(* IEC 61131-3 sources: daoli-st-library/_quarantine/R80, 3 files *)

(* ---- FC_DL_HydroPipePressDrop.st ---- *)
(*
  ============================================================
  组件名 : FC_DL_HydroPipePressDrop
  分类   : DL_Device
  功能   : 液压管路压降计算，由流量管径长度求流速、雷诺数、摩阻系数与压降
  开源溯源 : internal-design（本轮无外部代码逐行引用）
             参考语义 : 无外部参考
  复杂度 : C2
  版本   : 1.0.0
  ============================================================
  口径说明 : 工作介质取液压油，密度按 850 kg/m3 常量代入；黏度由 cSt 折算为 m2/s；
             层流区用 64/Re，湍流区用 Blasius 式 0.3164/Re^0.25；粗糙度引脚仅登记
             供上层记录，本件不进入摩阻判据（Colebrook 迭代属另一件边界）。
*)

FUNCTION FC_DL_HydroPipePressDrop : REAL
VAR_INPUT
    rFlow_lpm  : REAL; // 体积流量 [l/min] volume flow [l per minute]
    rDia_mm    : REAL; // 管内径 [mm] pipe inner diameter [mm]
    rLength_m  : REAL; // 管长 [m] pipe length [m]
    rVisc_cSt  : REAL; // 运动黏度 [cSt] kinematic viscosity [centistoke]
    rRough_mm  : REAL; // 管内壁粗糙度 [mm] inner wall roughness [mm]
END_VAR
VAR_OUTPUT
    rVel_m_s : REAL; // 管内流速 [m/s] pipe velocity [m per second]
    rRe      : REAL; // 雷诺数 [无量纲] Reynolds number [dimensionless]
    rDrop_bar: REAL; // 沿程压降 [bar] friction pressure drop [bar]
    bValid   : BOOL; // 结果有效标志 result validity flag
END_VAR
VAR CONSTANT
    DL_PI_4     : REAL := 0.7853982; // 四分之圆周率 pi divided by four
    DL_MM_TO_M  : REAL := 1000.0; // 每米毫米数 millimetres per metre
    DL_LPM_TO_M3S : REAL := 60000.0; // 升每分到立方米每秒的除数 divisor from litre per minute to cubic metre per second
    DL_CST_TO_M2S : REAL := 1.0E-6; // 厘斯到平方米每秒的乘子 multiplier from centistoke to square metre per second
    DL_DENSITY  : REAL := 850.0; // 液压油密度 [kg/m3] hydraulic oil density [kg per cubic metre]
    DL_RE_LAM   : REAL := 2300.0; // 层流上限雷诺数 laminar Reynolds ceiling
    DL_LAM_COEF : REAL := 64.0; // 层流摩阻系数分子 laminar friction numerator
    DL_BLA_COEF : REAL := 0.3164; // Blasius 式系数 Blasius coefficient
    DL_BLA_EXP  : REAL := 0.25; // Blasius 式指数 Blasius exponent
    DL_PA_TO_BAR: REAL := 100000.0; // 帕到巴换算 pascal per bar
END_VAR
VAR
    _bFin  : BOOL := FALSE; // 五输入有限性判定 finiteness verdict of the five inputs
    _rDiaM : REAL := 0.0; // 管径折算 [m] diameter in metre [m]
    _rArea : REAL := 0.0; // 管截面面积 [m2] pipe section area [m2]
    _rNu   : REAL := 0.0; // 运动黏度折算 [m2/s] viscosity in square metre per second
    _rQ    : REAL := 0.0; // 体积流量折算 [m3/s] flow in cubic metre per second
    _rVel  : REAL := 0.0; // 流速中间量 [m/s] intermediate velocity [m per second]
    _rRe   : REAL := 0.0; // 雷诺数中间量 [无量纲] intermediate Reynolds number [dimensionless]
    _rLam  : REAL := 0.0; // 摩阻系数 [无量纲] friction factor [dimensionless]
    _rDrop : REAL := 0.0; // 压降中间量 [Pa] intermediate drop [pascal]
END_VAR

// 段 1｜出口预置 preset the exit
FC_DL_HydroPipePressDrop := 0.0; // 缺省返回零 default zero return
rVel_m_s := 0.0; // 流速预置零 velocity preset to zero
rRe := 0.0; // 雷诺数预置零 Reynolds preset to zero
rDrop_bar := 0.0; // 压降预置零 drop preset to zero
bValid := FALSE; // 计算完成前不认结果 unusable before the calculation
// 段 2｜非有限闸 finiteness gate
_bFin := (rFlow_lpm = rFlow_lpm) AND (rDia_mm = rDia_mm) AND (rLength_m = rLength_m) AND (rVisc_cSt = rVisc_cSt) AND (rRough_mm = rRough_mm); // 五输入自反判定 self comparison of the five inputs
IF NOT _bFin THEN
    RETURN; // 非有限即无效 non finite means invalid
END_IF
// 段 3｜几何与黏度闸 geometry and viscosity gate
IF (rDia_mm <= 0.0) OR (rLength_m < 0.0) OR (rFlow_lpm < 0.0) THEN
    RETURN; // 管径非正或负长度负流量 an illegal diameter length or flow
END_IF
IF rVisc_cSt <= 0.0 THEN
    RETURN; // 黏度非正无法算雷诺数 a non positive viscosity cannot carry Reynolds
END_IF
// 段 4｜流速与雷诺数 velocity and the Reynolds number
_rDiaM := rDia_mm / DL_MM_TO_M; // 管径折算为米 convert the diameter to metre
_rArea := DL_PI_4 * _rDiaM * _rDiaM; // 管截面面积 pipe section area
_rQ := rFlow_lpm / DL_LPM_TO_M3S; // 流量折算为立方米每秒 convert the flow
_rVel := _rQ / _rArea; // 流速，除子为已证正面积 velocity over a proven positive area
_rNu := rVisc_cSt * DL_CST_TO_M2S; // 黏度折算为平方米每秒 convert the viscosity
_rRe := _rVel * _rDiaM / _rNu; // 雷诺数，除子为已证正黏度 Reynolds over a proven positive viscosity
rVel_m_s := _rVel; // 流速落定 land the velocity
rRe := _rRe; // 雷诺数落定 land the Reynolds number
// 段 5｜零流早退：雷诺数近零时压降为零 zero flow early exit with a zero drop
IF _rRe < 1.0 THEN
    bValid := TRUE; // 零流工况结果有效 a zero flow case is still usable
    RETURN; // 压降保持零 the drop stays zero
END_IF
// 段 6｜摩阻系数分区分支 friction factor by flow regime
IF _rRe < DL_RE_LAM THEN
    _rLam := DL_LAM_COEF / _rRe; // 层流区 sixty four over Reynolds
ELSE
    IF _rRe > 1.0E30 THEN
        RETURN; // 雷诺数越出数值上限 refuse an out of scale Reynolds number
    END_IF
    _rLam := DL_BLA_COEF / EXPT(_rRe, DL_BLA_EXP); // 湍流区 Blasius 式 the Blasius form for the turbulent regime
END_IF
// 段 7｜压降与出口 drop and the exit
_rDrop := _rLam * (rLength_m / _rDiaM) * (DL_DENSITY * _rVel * _rVel / 2.0); // 沿程压降 friction pressure drop
rDrop_bar := _rDrop / DL_PA_TO_BAR; // 压降换算为巴 convert the drop to bar
bValid := TRUE; // 结果可用 result usable
FC_DL_HydroPipePressDrop := rDrop_bar; // 函数返回压降 return the drop
END_FUNCTION

(* ---- FC_DL_StatsGeoMeanCalc.st ---- *)
(*
  ============================================================
  组件名 : FC_DL_StatsGeoMeanCalc
  分类   : DL_MathData
  功能   : 定长样本的几何平均值计算，非正值剔除后按自然对数均值再取指数
  开源溯源 : internal-design（本轮无外部代码逐行引用）
             参考语义 : 无外部参考
  复杂度 : C1
  版本   : 1.0.0
  ============================================================
*)

FUNCTION FC_DL_StatsGeoMeanCalc : REAL
VAR_INPUT
    aData  : ARRAY[0..31] OF REAL; // 样本数组，定长三十二 [工程单位] sample array of thirty two fixed slots [engineering unit]
    nCount : INT; // 有效样本数 1~32 [个] effective sample count from one to thirty two [count]
    rMinPos: REAL; // 正样本下限，非正或非有限时回默认值 [工程单位] positive sample floor, non positive values fall back to the default [engineering unit]
END_VAR
VAR_OUTPUT
    rGeoMean : REAL; // 几何平均值 [工程单位] geometric mean [engineering unit]
    nSkipped : INT; // 被剔除的样本数 [个] skipped sample count [count]
    bValid   : BOOL; // 结果有效标志 result validity flag
END_VAR
VAR CONSTANT
    DL_CAP  : INT := 32; // 数组容量 [个] array capacity [count]
    DL_POS_FLOOR : REAL := 1.0E-9; // 正样本下限默认值 default positive sample floor
END_VAR
VAR
    i      : INT := 0; // 遍历游标 [个] walk cursor [count]
    nOk    : INT := 0; // 参与取对数的样本数 [个] sample count entering the logarithm [count]
    _rSumLn: REAL := 0.0; // 自然对数和 [无量纲] sum of natural logarithms [dimensionless]
    _rFloor: REAL := 0.0; // 钳位后的正样本下限 [工程单位] clamped positive sample floor [engineering unit]
    _rGeo  : REAL := 0.0; // 几何均值中间量 [工程单位] intermediate geometric mean [engineering unit]
END_VAR

// 段 1｜出口预置 preset the exit
FC_DL_StatsGeoMeanCalc := 0.0; // 缺省返回零 default zero return
rGeoMean := 0.0; // 几何均值预置零 geometric mean preset to zero
nSkipped := 0; // 剔除数预置零 skipped count preset to zero
bValid := FALSE; // 计算完成前不认结果 unusable before the calculation
// 段 2｜点数闸与下限整形 count gate and floor reshape
IF (nCount < 1) OR (nCount > DL_CAP) THEN
    RETURN; // 点数越界即无效 an out of range count is void
END_IF
_rFloor := rMinPos; // 取入参正样本下限 take the positive floor input
IF _rFloor <> _rFloor THEN
    _rFloor := DL_POS_FLOOR; // 非有限下限回默认值 a non finite floor falls back to the default
ELSIF _rFloor <= 0.0 THEN
    _rFloor := DL_POS_FLOOR; // 非正下限回默认值 a non positive floor falls back to the default
END_IF
// 段 3｜剔除与对数累加 skip the ineligible samples and accumulate logarithms
FOR i := 0 TO (nCount - 1) DO
    IF (aData[i] <> aData[i]) OR (aData[i] < _rFloor) THEN
        nSkipped := nSkipped + 1; // 非有限或非正样本剔除 skip a non finite or a non positive sample
    ELSE
        _rSumLn := _rSumLn + LN(aData[i]); // 自然对数累加 accumulate the natural logarithm
        nOk := nOk + 1; // 有效样本计数 count the usable sample
    END_IF
END_FOR
// 段 4｜全剔除闸 the all skipped gate
IF nOk <= 0 THEN
    RETURN; // 无正样本时几何均值无定义 an all skipped set has no geometric mean
END_IF
// 段 5｜指数还原与出口 exponent restore and the exit
_rGeo := EXP(_rSumLn / INT_TO_REAL(nOk)); // 对数均值取指数，除子为已证正计数 exponent of the mean logarithm
IF (_rGeo <> _rGeo) OR (ABS(_rGeo) > 1.0E30) THEN
    RETURN; // 结果非有限拒收 refuse a non finite result
END_IF
rGeoMean := _rGeo; // 几何均值落定 land the geometric mean
bValid := TRUE; // 结果可用 result usable
FC_DL_StatsGeoMeanCalc := _rGeo; // 函数返回几何均值 return the geometric mean
END_FUNCTION

(* ---- FC_DL_StatsIqrCalc.st ---- *)
(*
  ============================================================
  组件名 : FC_DL_StatsIqrCalc
  分类   : DL_MathData
  功能   : 定长样本的四分位距与异常栅栏计算，先插入排序再按位置线性插值
  开源溯源 : internal-design（本轮无外部代码逐行引用）
             参考语义 : 无外部参考
  复杂度 : C2
  版本   : 1.0.0
  ============================================================
  口径说明 : 分位位置取 (n-1) 法，Q1 位置 0.25×(n-1)、Q3 位置 0.75×(n-1)，
             位置非整数时按相邻两个样本线性插值；栅栏取 Q1-1.5×IQR 与 Q3+1.5×IQR。
             样本数小于二时四分位无定义，本件判无效。
*)

FUNCTION FC_DL_StatsIqrCalc : REAL
VAR_INPUT
    aData  : ARRAY[0..31] OF REAL; // 样本数组，定长三十二 [工程单位] sample array of thirty two fixed slots [engineering unit]
    nCount : INT; // 有效样本数 2~32 [个] effective sample count from two to thirty two [count]
END_VAR
VAR_OUTPUT
    rQ1        : REAL; // 下四分位 [工程单位] lower quartile [engineering unit]
    rQ3        : REAL; // 上四分位 [工程单位] upper quartile [engineering unit]
    rIqr       : REAL; // 四分位距 [工程单位] interquartile range [engineering unit]
    rFenceLow  : REAL; // 下栅栏 [工程单位] lower fence [engineering unit]
    rFenceHigh : REAL; // 上栅栏 [工程单位] upper fence [engineering unit]
    bValid     : BOOL; // 结果有效标志 result validity flag
END_VAR
VAR CONSTANT
    DL_CAP   : INT := 32; // 数组容量 [个] array capacity [count]
    DL_Q1    : REAL := 0.25; // 下四分位位置系数 lower quartile position factor
    DL_Q3    : REAL := 0.75; // 上四分位位置系数 upper quartile position factor
    DL_FENCE : REAL := 1.5; // 栅栏系数 fence factor
END_VAR
VAR
    aBuf  : ARRAY[0..31] OF REAL; // 排序副本 [工程单位] sorted copy [engineering unit]
    i     : INT := 0; // 外层游标 [个] outer cursor [count]
    j     : INT := 0; // 内层游标 [个] inner cursor [count]
    nIdx  : INT := 0; // 插值左邻下标 [个] left neighbour index [count]
    _rKey : REAL := 0.0; // 插入排序待插值 [工程单位] insertion key [engineering unit]
    _rPos : REAL := 0.0; // 分位位置 [位] quantile position [slot]
    _rFrac: REAL := 0.0; // 位置小数部分 [无量纲] fractional part of the position [dimensionless]
    _rQ1  : REAL := 0.0; // 下四分位中间量 [工程单位] intermediate lower quartile [engineering unit]
    _rQ3  : REAL := 0.0; // 上四分位中间量 [工程单位] intermediate upper quartile [engineering unit]
END_VAR

// 段 1｜出口预置 preset the exit
FC_DL_StatsIqrCalc := 0.0; // 缺省返回零 default zero return
rQ1 := 0.0; // 下四分位预置零 lower quartile preset to zero
rQ3 := 0.0; // 上四分位预置零 upper quartile preset to zero
rIqr := 0.0; // 四分位距预置零 interquartile range preset to zero
rFenceLow := 0.0; // 下栅栏预置零 lower fence preset to zero
rFenceHigh := 0.0; // 上栅栏预置零 upper fence preset to zero
bValid := FALSE; // 计算完成前不认结果 unusable before the calculation
// 段 2｜点数闸 sample count gate
IF (nCount < 2) OR (nCount > DL_CAP) THEN
    RETURN; // 点数越界或不足二即无效 an out of range or a too small count is void
END_IF
// 段 3｜拷贝并插入排序 copy then insertion sort
FOR i := 0 TO (nCount - 1) DO
    IF aData[i] <> aData[i] THEN
        RETURN; // 非有限样本拒收，出口保持零点 refuse a non finite sample
    END_IF
    aBuf[i] := aData[i]; // 逐点拷贝 copy sample by sample
END_FOR
FOR i := 1 TO (nCount - 1) DO
    _rKey := aBuf[i]; // 待插值取当前点 the key is the current sample
    j := i - 1; // 内层游标从左邻起 the inner cursor starts at the left neighbour
    WHILE (j >= 0) AND (aBuf[j] > _rKey) DO
        aBuf[j + 1] := aBuf[j]; // 后移空位 shift right to open a slot
        j := j - 1; // 游标左退 step the cursor left
    END_WHILE
    aBuf[j + 1] := _rKey; // 落位 drop the key in place
END_FOR
// 段 4｜下四分位插值 lower quartile interpolation
_rPos := DL_Q1 * INT_TO_REAL(nCount - 1); // 下四分位位置 lower quartile position
nIdx := REAL_TO_INT(FLOOR(_rPos)); // 左邻下标，先向下取整再转整型 floor then convert to integer
IF nIdx > (nCount - 2) THEN
    nIdx := nCount - 2; // 左邻下标钳位 clamp the left neighbour index
END_IF
_rFrac := _rPos - INT_TO_REAL(nIdx); // 位置小数部分 fractional part of the position
_rQ1 := aBuf[nIdx] + _rFrac * (aBuf[nIdx + 1] - aBuf[nIdx]); // 相邻样本线性插值 linear blend of the neighbours
// 段 5｜上四分位插值 upper quartile interpolation
_rPos := DL_Q3 * INT_TO_REAL(nCount - 1); // 上四分位位置 upper quartile position
nIdx := REAL_TO_INT(FLOOR(_rPos)); // 左邻下标，先向下取整再转整型 floor then convert to integer
IF nIdx > (nCount - 2) THEN
    nIdx := nCount - 2; // 左邻下标钳位 clamp the left neighbour index
END_IF
_rFrac := _rPos - INT_TO_REAL(nIdx); // 位置小数部分 fractional part of the position
_rQ3 := aBuf[nIdx] + _rFrac * (aBuf[nIdx + 1] - aBuf[nIdx]); // 相邻样本线性插值 linear blend of the neighbours
// 段 6｜四分位距与栅栏 interquartile range and the fences
rQ1 := _rQ1; // 下四分位落定 land the lower quartile
rQ3 := _rQ3; // 上四分位落定 land the upper quartile
rIqr := _rQ3 - _rQ1; // 四分位距 interquartile range
rFenceLow := _rQ1 - DL_FENCE * rIqr; // 下栅栏 lower fence
rFenceHigh := _rQ3 + DL_FENCE * rIqr; // 上栅栏 upper fence
bValid := TRUE; // 结果可用 result usable
FC_DL_StatsIqrCalc := rIqr; // 函数返回四分位距 return the range
END_FUNCTION
